Staubli VAL3: cycle_Stop.pgx

program cycle_Stop()
begin
  //进程:Stopping
  rs:_nOmacStat=8
  // Stop task
  taskKill("Reset")
  taskKill("Start")
  taskKill("productCycle")
  taskKill("End")
  taskKill("GoHome")
  taskKill("Monitor")
  taskKill("RotGoHome")
  taskKill("Monitor1")
  taskKill("getForce")

  while !isPowered()
    enablePower()
    delay(1)
  endWhile
  //
  stopMove()
  call ar:getCurMoveID(bGetMovId,"Stop")
  resetMotion()
  disablePower()
  wait(isPowered()==false)
  //2025.7.21 add 复位输出信号
  call plc:resetOutput()
  //OMAC进程:Stopped
  rs:_nOmacStat=9
  logMsg("当前处于生产停止状态 "+toString(".2",clock()))
  rs:_sRobotStatus="当前处于生产停止状态"
  delay(0)
end
